// Nombre → état de calibration (restauration) ; une calibration en cours à la sauvegarde revient « jamais faite »
FUNCTION F_CalibStateOf : E_CalibState
VAR_INPUT
    fValue : LREAL;
END_VAR

IF fValue > 2.5 AND fValue < 3.5 THEN
    F_CalibStateOf := E_CalibState.Failed;
ELSIF fValue > 1.5 AND fValue < 2.5 THEN
    F_CalibStateOf := E_CalibState.Expired;
ELSIF fValue > 0.5 AND fValue < 1.5 THEN
    F_CalibStateOf := E_CalibState.Valid;
ELSE
    F_CalibStateOf := E_CalibState.Never;
END_IF

END_FUNCTION

(* stored: Version 1.1.0.1, ProductVersion 3.1.4024.12
   POU F_CalibStateOf: Id {298b929f-60ee-5b92-bf51-cd05cbb89e95}, SpecialFunc None *)
